// TIA Portal V21 export
// export: Created 2026-08-21T20:18:52.4495075Z, ExportSetting None, DisplayName Totally Integrated Automation Portal, DisplayVersion V21, DisplayName STEP 7 Professional, DisplayVersion V21, DisplayName STEP 7 Safety, DisplayVersion V21, DisplayName Tech WebApplication, DisplayVersion V21, DisplayName WinCC Basic/Comfort/Advanced, DisplayVersion V21, DisplayName WinCC Professional, DisplayVersion V21, DisplayName WinCC Unified, DisplayVersion V21
DATA_BLOCK "Service_Interaction_FB_DB"   // DB57
// stored: InstanceOfName Service_Interaction_FB, InstanceOfType FB
"Service_Interaction_FB"
   // VAR_INPUT
   //    Startbit { ExternalAccessible := 'False'; ExternalVisible := 'False'; ExternalWritable := 'False'} : Bool;
   //    AnswerID { ExternalAccessible := 'False'; ExternalVisible := 'False'; ExternalWritable := 'False'} : DWord;
   // END_VAR
   // VAR_OUTPUT
   //    P100_Start : Bool;
   //    P101_Start : Bool;
   // END_VAR
   // VAR_IN_OUT
   //    Pump_100 : "MotL";
   //    Pump_101 : "MotL";
   // END_VAR
BEGIN
END_DATA_BLOCK
